Fanuc KAREL source: kd00051.KL

PROGRAM KD00051
%STACKSIZE=65535
%PRIORITY=65535
%NOLOCKGROUP
VAR
I : INTEGER
J : INTEGER
B : BOOLEAN
R : REAL
S : STRING[80]
P : POSITION
BEGIN
-- UNRESOLVED_PC line 12 opcodes [01 22 1C 2E 0A 82 0B] marker_code=0
END KD00051
